Staubli VAL3: resfreshTRAJ.pgx

program resfreshTRAJ(string x_sHtml)
  local num l_nSize
  local num l_nSize1
  local num l_i
begin
  call trajectory:getSize(l_nSize)
  call trajectory:getTrajList(sTRAJList)

  if l_nSize>49
    nPgNumPROG=roundUp(l_nSize/49)
  else
    nPgNumPROG=1
  endIf

  l_nSize1=l_nSize%49

  if nPgIndexPROG==nPgNumPROG-1
    if l_nSize1!=0
      resize(sList,1,l_nSize1)
      for l_i = 0 to size(sList)-1
        sList[l_i]=sTRAJList[l_i+nPgIndexPROG*49]
      endFor
    else
      resize(sList,1,49)
      for l_i = 0 to size(sList)-1
        sList[l_i]=sTRAJList[l_i+nPgIndexPROG*49]
      endFor
    endIf
  else
    resize(sList,1,49)
    for l_i = 0 to size(sList)-1
      sList[l_i]=sTRAJList[l_i+nPgIndexPROG*49]
    endFor
  endIf
  userPageBind(x_sHtml,"lst1","options",sList,size(sList),"r")
  sPagePROG=toString("",nPgNumPROG)
  sPgIndexPROG=toString("",nPgIndexPROG+1)
end
